(* PLC project ldtest *)

PROGRAM LdDemo

(* LD diagram, written out as Structured Text *)
%QX0.0 := (%IX0.0 OR %IX0.1) AND NOT %IX0.2;
END_PROGRAM
